Fanuc KAREL source: KA00074.KL

PROGRAM KA00074
%NOLOCKGROUP
VAR
  SRC: XYZWPREXT
  DST: REAL
BEGIN
  SRC.X = 1.0
  DST = SRC
END KA00074
